(* IEC 61131-3 sources: Jacob-Formschaumtechnik-ISEL-CNC-Retrofit/twincat/PLC/src/7_Weitere, 1 file *)

(* ---- MAIN.st ---- *)
PROGRAM MAIN
VAR
END_VAR

PRG_Test();   (* Simulationstest, nur aktiv mit bTestEnable im Simulations-Build *)
PRG_Main();
END_PROGRAM
